TYPE ST_EL6633 :
STRUCT
	sTerminalName : STRING(80) := 'EL6633 | 2-Port PROFINET Communication Interface';

    stTerminalInfo : ST_Terminal_Info;
END_STRUCT
END_TYPE

(* stored: Version 1.1.0.1, ProductVersion 3.1.4026.18
   DUT ST_EL6633: Id {9a411c2d-88d5-49e1-bdd7-f4a2b00ecdd0} *)
